    PROC Path_ContornoExterno()
        MoveJ Pivote,v100,z1,MyNewTool\WObj:=Cara;
        MoveJ Target_190,v100,z1,MyNewTool\WObj:=Cara;
        MoveL Target_200,v100,z1,MyNewTool\WObj:=Cara;
        MoveL Target_210,v100,z1,MyNewTool\WObj:=Cara;
        MoveL Target_220,v100,z1,MyNewTool\WObj:=Cara;
        MoveL Target_230,v100,z1,MyNewTool\WObj:=Cara;
        MoveL Target_240,v100,z1,MyNewTool\WObj:=Cara;
        MoveL Target_250,v100,z1,MyNewTool\WObj:=Cara;
        MoveL Target_260,v100,z1,MyNewTool\WObj:=Cara;
        MoveL Target_270,v100,z1,MyNewTool\WObj:=Cara;
        MoveL Target_280,v100,z1,MyNewTool\WObj:=Cara;
        MoveL Target_290,v100,z1,MyNewTool\WObj:=Cara;
        MoveL Target_300,v100,z1,MyNewTool\WObj:=Cara;
        MoveL Target_310,v100,z1,MyNewTool\WObj:=Cara;
        MoveL Target_320,v100,z1,MyNewTool\WObj:=Cara;
        MoveL Target_330,v100,z1,MyNewTool\WObj:=Cara;
        MoveL Target_340,v100,z1,MyNewTool\WObj:=Cara;
        MoveL Target_350,v100,z1,MyNewTool\WObj:=Cara;
        MoveL Target_360,v100,z1,MyNewTool\WObj:=Cara;
        MoveL Target_370,v100,z1,MyNewTool\WObj:=Cara;
        MoveL Target_380,v100,z1,MyNewTool\WObj:=Cara;
        MoveL Target_390,v100,z1,MyNewTool\WObj:=Cara;
        MoveL Target_400,v100,z1,MyNewTool\WObj:=Cara;
        MoveL Target_410,v100,z1,MyNewTool\WObj:=Cara;
        MoveL Target_420,v100,z1,MyNewTool\WObj:=Cara;
        MoveL Target_430,v100,z1,MyNewTool\WObj:=Cara;
        MoveL Target_440,v100,z1,MyNewTool\WObj:=Cara;
        MoveL Target_450,v100,z1,MyNewTool\WObj:=Cara;
        MoveL Target_460,v100,z1,MyNewTool\WObj:=Cara;
        MoveL Target_470,v100,z1,MyNewTool\WObj:=Cara;
        MoveL Target_480,v100,z1,MyNewTool\WObj:=Cara;
        MoveL Target_490,v100,z1,MyNewTool\WObj:=Cara;
        MoveL Target_500,v100,z1,MyNewTool\WObj:=Cara;
        MoveL Target_510,v100,z1,MyNewTool\WObj:=Cara;
        MoveL Target_520,v100,z1,MyNewTool\WObj:=Cara;
        MoveL Target_530,v100,z1,MyNewTool\WObj:=Cara;
        MoveL Target_540,v100,z1,MyNewTool\WObj:=Cara;
        MoveL Target_550,v100,z1,MyNewTool\WObj:=Cara;
        MoveL Target_560,v100,z1,MyNewTool\WObj:=Cara;
        MoveL Target_570,v100,z1,MyNewTool\WObj:=Cara;
        MoveL Target_580,v100,z1,MyNewTool\WObj:=Cara;
        MoveL Target_590,v100,z1,MyNewTool\WObj:=Cara;
        MoveL Target_600,v100,z1,MyNewTool\WObj:=Cara;
        MoveL Target_610,v100,z1,MyNewTool\WObj:=Cara;
        MoveL Target_620,v100,z1,MyNewTool\WObj:=Cara;
        MoveL Target_630,v100,z1,MyNewTool\WObj:=Cara;
        MoveL Target_640,v100,z1,MyNewTool\WObj:=Cara;
        MoveL Target_650,v100,z1,MyNewTool\WObj:=Cara;
        MoveL Target_660,v100,z1,MyNewTool\WObj:=Cara;
        MoveL Target_670,v100,z1,MyNewTool\WObj:=Cara;
        MoveL Target_680,v100,z1,MyNewTool\WObj:=Cara;
        MoveL Target_690,v100,z1,MyNewTool\WObj:=Cara;
        MoveL Target_700,v100,z1,MyNewTool\WObj:=Cara;
        MoveL Target_710,v100,z1,MyNewTool\WObj:=Cara;
        MoveL Target_720,v100,z1,MyNewTool\WObj:=Cara;
        MoveL Target_730,v100,z1,MyNewTool\WObj:=Cara;
        MoveL Target_740,v100,z1,MyNewTool\WObj:=Cara;
        MoveL Target_750,v100,z1,MyNewTool\WObj:=Cara;
        MoveL Target_760,v100,z1,MyNewTool\WObj:=Cara;
        MoveL Target_770,v100,z1,MyNewTool\WObj:=Cara;
        MoveL Target_780,v100,z1,MyNewTool\WObj:=Cara;
        MoveL Target_790,v100,z1,MyNewTool\WObj:=Cara;
        MoveL Target_800,v100,z1,MyNewTool\WObj:=Cara;
        MoveL Target_810,v100,z1,MyNewTool\WObj:=Cara;
        MoveL Target_820,v100,z1,MyNewTool\WObj:=Cara;
        MoveL Target_830,v100,z1,MyNewTool\WObj:=Cara;
        MoveL Target_840,v100,z1,MyNewTool\WObj:=Cara;
        MoveL Target_850,v100,z1,MyNewTool\WObj:=Cara;
        MoveL Target_860,v100,z1,MyNewTool\WObj:=Cara;
        MoveL Target_870,v100,z1,MyNewTool\WObj:=Cara;
        MoveL Target_880,v100,z1,MyNewTool\WObj:=Cara;
        MoveL Target_890,v100,z1,MyNewTool\WObj:=Cara;
        MoveL Target_900,v100,z1,MyNewTool\WObj:=Cara;
        MoveL Target_910,v100,z1,MyNewTool\WObj:=Cara;
        MoveL Target_920,v100,z1,MyNewTool\WObj:=Cara;
        MoveL Target_930,v100,z1,MyNewTool\WObj:=Cara;
        MoveL Target_940,v100,z1,MyNewTool\WObj:=Cara;
        MoveL Target_950,v100,z1,MyNewTool\WObj:=Cara;
        MoveL Target_960,v100,z1,MyNewTool\WObj:=Cara;
        MoveL Target_970,v100,z1,MyNewTool\WObj:=Cara;
        MoveL Target_980,v100,z1,MyNewTool\WObj:=Cara;
        MoveL Target_990,v100,z1,MyNewTool\WObj:=Cara;
        MoveL Target_1000,v100,z1,MyNewTool\WObj:=Cara;
        MoveL Target_1010,v100,z1,MyNewTool\WObj:=Cara;
        MoveL Target_1020,v100,z1,MyNewTool\WObj:=Cara;
        MoveL Target_1030,v100,z1,MyNewTool\WObj:=Cara;
        MoveL Target_1040,v100,z1,MyNewTool\WObj:=Cara;
        MoveL Target_1050,v100,z1,MyNewTool\WObj:=Cara;
        MoveL Target_1060,v100,z1,MyNewTool\WObj:=Cara;
        MoveL Target_1070,v100,z1,MyNewTool\WObj:=Cara;
        MoveL Target_1080,v100,z1,MyNewTool\WObj:=Cara;
        MoveL Target_1090,v100,z1,MyNewTool\WObj:=Cara;
        MoveL Target_1100,v100,z1,MyNewTool\WObj:=Cara;
        MoveL Target_1110,v100,z1,MyNewTool\WObj:=Cara;
        MoveL Target_1120,v100,z1,MyNewTool\WObj:=Cara;
        MoveL Target_1130,v100,z1,MyNewTool\WObj:=Cara;
        MoveL Target_1140,v100,z1,MyNewTool\WObj:=Cara;
        MoveL Target_1150,v100,z1,MyNewTool\WObj:=Cara;
        MoveL Target_1160,v100,z1,MyNewTool\WObj:=Cara;
        MoveL Target_1170,v100,z1,MyNewTool\WObj:=Cara;
    ENDPROC
    PROC Path_Cabello()
        MoveJ Target_1350,v100,z1,MyNewTool\WObj:=Cara;
        MoveL Target_1360,v100,z1,MyNewTool\WObj:=Cara;
        MoveL Target_1370,v100,z1,MyNewTool\WObj:=Cara;
        MoveL Target_1380,v100,z1,MyNewTool\WObj:=Cara;
        MoveL Target_1390,v100,z1,MyNewTool\WObj:=Cara;
        MoveL Target_1400,v100,z1,MyNewTool\WObj:=Cara;
        MoveL Target_1410,v100,z1,MyNewTool\WObj:=Cara;
        MoveL Target_1420,v100,z1,MyNewTool\WObj:=Cara;
        MoveL Target_1430,v100,z1,MyNewTool\WObj:=Cara;
        MoveL Target_1440,v100,z1,MyNewTool\WObj:=Cara;
        MoveL Target_1450,v100,z1,MyNewTool\WObj:=Cara;
        MoveL Target_1460,v100,z1,MyNewTool\WObj:=Cara;
        MoveL Target_1470,v100,z1,MyNewTool\WObj:=Cara;
        MoveL Target_1480,v100,z1,MyNewTool\WObj:=Cara;
        MoveL Target_1490,v100,z1,MyNewTool\WObj:=Cara;
        MoveL Target_1500,v100,z1,MyNewTool\WObj:=Cara;
        MoveL Target_1510,v100,z1,MyNewTool\WObj:=Cara;
        MoveL Target_1520,v100,z1,MyNewTool\WObj:=Cara;
        MoveL Target_1530,v100,z1,MyNewTool\WObj:=Cara;
        MoveL Target_1540,v100,z1,MyNewTool\WObj:=Cara;
        MoveL Target_1550,v100,z1,MyNewTool\WObj:=Cara;
        MoveL Target_1560,v100,z1,MyNewTool\WObj:=Cara;
        MoveL Target_1570,v100,z1,MyNewTool\WObj:=Cara;
        MoveL Target_1580,v100,z1,MyNewTool\WObj:=Cara;
        MoveL Target_1590,v100,z1,MyNewTool\WObj:=Cara;
        MoveL Target_1600,v100,z1,MyNewTool\WObj:=Cara;
        MoveL Target_1610,v100,z1,MyNewTool\WObj:=Cara;
        MoveL Target_1620,v100,z1,MyNewTool\WObj:=Cara;
        MoveL Target_1630,v100,z1,MyNewTool\WObj:=Cara;
        MoveL Target_1640,v100,z1,MyNewTool\WObj:=Cara;
        MoveL Target_1650,v100,z1,MyNewTool\WObj:=Cara;
        MoveL Target_1660,v100,z1,MyNewTool\WObj:=Cara;
        MoveL Target_1670,v100,z1,MyNewTool\WObj:=Cara;
        MoveL Target_1680,v100,z1,MyNewTool\WObj:=Cara;
        MoveL Target_1690,v100,z1,MyNewTool\WObj:=Cara;
        MoveL Target_1700,v100,z1,MyNewTool\WObj:=Cara;
        MoveL Target_1710,v100,z1,MyNewTool\WObj:=Cara;
        MoveL Target_1720,v100,z1,MyNewTool\WObj:=Cara;
        MoveL Target_1730,v100,z1,MyNewTool\WObj:=Cara;
        MoveL Target_1740,v100,z1,MyNewTool\WObj:=Cara;
        MoveL Target_1750,v100,z1,MyNewTool\WObj:=Cara;
        MoveL Target_1760,v100,z1,MyNewTool\WObj:=Cara;
        MoveL Target_1770,v100,z1,MyNewTool\WObj:=Cara;
        MoveL Target_1780,v100,z1,MyNewTool\WObj:=Cara;
        MoveL Target_1790,v100,z1,MyNewTool\WObj:=Cara;
        MoveL Target_1800,v100,z1,MyNewTool\WObj:=Cara;
        MoveL Target_1810,v100,z1,MyNewTool\WObj:=Cara;
        MoveL Target_1820,v100,z1,MyNewTool\WObj:=Cara;
        MoveL Target_1830,v100,z1,MyNewTool\WObj:=Cara;
        MoveL Target_1840,v100,z1,MyNewTool\WObj:=Cara;
        MoveL Target_1850,v100,z1,MyNewTool\WObj:=Cara;
        MoveL Target_1860,v100,z1,MyNewTool\WObj:=Cara;
        MoveL Target_1870,v100,z1,MyNewTool\WObj:=Cara;
        MoveL Target_1880,v100,z1,MyNewTool\WObj:=Cara;
        MoveL Target_1890,v100,z1,MyNewTool\WObj:=Cara;
        MoveL Target_1900,v100,z1,MyNewTool\WObj:=Cara;
        MoveL Target_1910,v100,z1,MyNewTool\WObj:=Cara;
        MoveL Target_1920,v100,z1,MyNewTool\WObj:=Cara;
        MoveL Target_1930,v100,z1,MyNewTool\WObj:=Cara;
        MoveL Target_1940,v100,z1,MyNewTool\WObj:=Cara;
        MoveL Target_1950,v100,z1,MyNewTool\WObj:=Cara;
        MoveL Target_1960,v100,z1,MyNewTool\WObj:=Cara;
        MoveL Target_1970,v100,z1,MyNewTool\WObj:=Cara;
        MoveL Target_1980,v100,z1,MyNewTool\WObj:=Cara;
        MoveL Target_1990,v100,z1,MyNewTool\WObj:=Cara;
        MoveL Target_2000,v100,z1,MyNewTool\WObj:=Cara;
        MoveL Target_2010,v100,z1,MyNewTool\WObj:=Cara;
        MoveL Target_2020,v100,z1,MyNewTool\WObj:=Cara;
        MoveL Target_2030,v100,z1,MyNewTool\WObj:=Cara;
        MoveL Target_2040,v100,z1,MyNewTool\WObj:=Cara;
        MoveL Target_2050,v100,z1,MyNewTool\WObj:=Cara;
        MoveL Target_2060,v100,z1,MyNewTool\WObj:=Cara;
        MoveL Target_2070,v100,z1,MyNewTool\WObj:=Cara;
        MoveL Target_2080,v100,z1,MyNewTool\WObj:=Cara;
        MoveL Target_2090,v100,z1,MyNewTool\WObj:=Cara;
        MoveL Target_2100,v100,z1,MyNewTool\WObj:=Cara;
        MoveL Target_2110,v100,z1,MyNewTool\WObj:=Cara;
        MoveL Target_2120,v100,z1,MyNewTool\WObj:=Cara;
        MoveL Target_2130,v100,z1,MyNewTool\WObj:=Cara;
        MoveL Target_2140,v100,z1,MyNewTool\WObj:=Cara;
        MoveL Target_2150,v100,z1,MyNewTool\WObj:=Cara;
    ENDPROC
    PROC Path_Frente()
        MoveJ Target_2430,v100,z1,MyNewTool\WObj:=Cara;
        MoveL Target_2440,v100,z1,MyNewTool\WObj:=Cara;
        MoveL Target_2450,v100,z1,MyNewTool\WObj:=Cara;
        MoveL Target_2460,v100,z1,MyNewTool\WObj:=Cara;
        MoveL Target_2470,v100,z1,MyNewTool\WObj:=Cara;
        MoveL Target_2480,v100,z1,MyNewTool\WObj:=Cara;
        MoveL Target_2490,v100,z1,MyNewTool\WObj:=Cara;
        MoveL Target_2500,v100,z1,MyNewTool\WObj:=Cara;
        MoveL Target_2510,v100,z1,MyNewTool\WObj:=Cara;
        MoveL Target_2520,v100,z1,MyNewTool\WObj:=Cara;
        MoveL Target_2530,v100,z1,MyNewTool\WObj:=Cara;
        MoveL Target_2540,v100,z1,MyNewTool\WObj:=Cara;
        MoveL Target_2550,v100,z1,MyNewTool\WObj:=Cara;
        MoveL Target_2560,v100,z1,MyNewTool\WObj:=Cara;
        MoveL Target_2570,v100,z1,MyNewTool\WObj:=Cara;
        MoveL Target_2580,v100,z1,MyNewTool\WObj:=Cara;
        MoveL Target_2590,v100,z1,MyNewTool\WObj:=Cara;
        MoveL Target_2600,v100,z1,MyNewTool\WObj:=Cara;
        MoveL Target_2610,v100,z1,MyNewTool\WObj:=Cara;
        MoveL Target_2620,v100,z1,MyNewTool\WObj:=Cara;
        MoveL Target_2630,v100,z1,MyNewTool\WObj:=Cara;
        MoveL Target_2640,v100,z1,MyNewTool\WObj:=Cara;
        MoveL Target_2650,v100,z1,MyNewTool\WObj:=Cara;
        MoveL Target_2660,v100,z1,MyNewTool\WObj:=Cara;
        MoveL Target_2670,v100,z1,MyNewTool\WObj:=Cara;
        MoveL Target_2680,v100,z1,MyNewTool\WObj:=Cara;
        MoveL Target_2690,v100,z1,MyNewTool\WObj:=Cara;
        MoveL Target_2700,v100,z1,MyNewTool\WObj:=Cara;
    ENDPROC
    PROC Path_ContornoCara()
        MoveJ Target_2710,v100,z1,MyNewTool\WObj:=Cara;
        MoveL Target_2720,v100,z1,MyNewTool\WObj:=Cara;
        MoveL Target_2730,v100,z1,MyNewTool\WObj:=Cara;
        MoveL Target_2740,v100,z1,MyNewTool\WObj:=Cara;
        MoveL Target_2750,v100,z1,MyNewTool\WObj:=Cara;
        MoveL Target_2760,v100,z1,MyNewTool\WObj:=Cara;
        MoveL Target_2770,v100,z1,MyNewTool\WObj:=Cara;
        MoveL Target_2780,v100,z1,MyNewTool\WObj:=Cara;
        MoveL Target_2790,v100,z1,MyNewTool\WObj:=Cara;
        MoveL Target_2800,v100,z1,MyNewTool\WObj:=Cara;
        MoveL Target_2810,v100,z1,MyNewTool\WObj:=Cara;
        MoveL Target_2820,v100,z1,MyNewTool\WObj:=Cara;
        MoveL Target_2830,v100,z1,MyNewTool\WObj:=Cara;
        MoveL Target_2840,v100,z1,MyNewTool\WObj:=Cara;
        MoveL Target_2850,v100,z1,MyNewTool\WObj:=Cara;
        MoveL Target_2860,v100,z1,MyNewTool\WObj:=Cara;
        MoveL Target_2870,v100,z1,MyNewTool\WObj:=Cara;
        MoveL Target_2880,v100,z1,MyNewTool\WObj:=Cara;
        MoveL Target_2890,v100,z1,MyNewTool\WObj:=Cara;
        MoveL Target_2900,v100,z1,MyNewTool\WObj:=Cara;
        MoveL Target_2910,v100,z1,MyNewTool\WObj:=Cara;
        MoveL Target_2920,v100,z1,MyNewTool\WObj:=Cara;
        MoveL Target_2930,v100,z1,MyNewTool\WObj:=Cara;
        MoveL Target_2940,v100,z1,MyNewTool\WObj:=Cara;
        MoveL Target_2950,v100,z1,MyNewTool\WObj:=Cara;
        MoveL Target_2960,v100,z1,MyNewTool\WObj:=Cara;
        MoveL Target_2970,v100,z1,MyNewTool\WObj:=Cara;
        MoveL Target_2980,v100,z1,MyNewTool\WObj:=Cara;
        MoveL Target_2990,v100,z1,MyNewTool\WObj:=Cara;
        MoveL Target_3000,v100,z1,MyNewTool\WObj:=Cara;
        MoveL Target_3010,v100,z1,MyNewTool\WObj:=Cara;
        MoveL Target_3020,v100,z1,MyNewTool\WObj:=Cara;
        MoveL Target_3030,v100,z1,MyNewTool\WObj:=Cara;
        MoveL Target_3040,v100,z1,MyNewTool\WObj:=Cara;
        MoveL Target_3050,v100,z1,MyNewTool\WObj:=Cara;
        MoveL Target_3060,v100,z1,MyNewTool\WObj:=Cara;
        MoveL Target_3070,v100,z1,MyNewTool\WObj:=Cara;
        MoveL Target_3080,v100,z1,MyNewTool\WObj:=Cara;
        MoveL Target_3090,v100,z1,MyNewTool\WObj:=Cara;
        MoveL Target_3100,v100,z1,MyNewTool\WObj:=Cara;
        MoveL Target_3110,v100,z1,MyNewTool\WObj:=Cara;
        MoveL Target_3120,v100,z1,MyNewTool\WObj:=Cara;
        MoveL Target_3130,v100,z1,MyNewTool\WObj:=Cara;
        MoveL Target_3140,v100,z1,MyNewTool\WObj:=Cara;
        MoveL Target_3150,v100,z1,MyNewTool\WObj:=Cara;
        MoveL Target_3160,v100,z1,MyNewTool\WObj:=Cara;
        MoveL Target_3170,v100,z1,MyNewTool\WObj:=Cara;
        MoveL Target_3180,v100,z1,MyNewTool\WObj:=Cara;
        MoveL Target_3190,v100,z1,MyNewTool\WObj:=Cara;
        MoveL Target_3200,v100,z1,MyNewTool\WObj:=Cara;
        MoveL Target_3210,v100,z1,MyNewTool\WObj:=Cara;
        MoveL Target_3220,v100,z1,MyNewTool\WObj:=Cara;
        MoveL Target_3230,v100,z1,MyNewTool\WObj:=Cara;
        MoveL Target_3240,v100,z1,MyNewTool\WObj:=Cara;
        MoveL Target_3250,v100,z1,MyNewTool\WObj:=Cara;
        MoveL Target_3260,v100,z1,MyNewTool\WObj:=Cara;
        MoveL Target_3270,v100,z1,MyNewTool\WObj:=Cara;
        MoveL Target_3280,v100,z1,MyNewTool\WObj:=Cara;
        MoveL Target_3290,v100,z1,MyNewTool\WObj:=Cara;
        MoveL Target_3300,v100,z1,MyNewTool\WObj:=Cara;
        MoveL Target_3310,v100,z1,MyNewTool\WObj:=Cara;
        MoveL Target_3320,v100,z1,MyNewTool\WObj:=Cara;
        MoveL Target_3330,v100,z1,MyNewTool\WObj:=Cara;
        MoveL Target_3340,v100,z1,MyNewTool\WObj:=Cara;
        MoveL Target_3350,v100,z1,MyNewTool\WObj:=Cara;
        MoveL Target_3360,v100,z1,MyNewTool\WObj:=Cara;
        MoveL Target_3370,v100,z1,MyNewTool\WObj:=Cara;
        MoveL Target_3380,v100,z1,MyNewTool\WObj:=Cara;
        MoveL Target_3390,v100,z1,MyNewTool\WObj:=Cara;
        MoveL Target_3400,v100,z1,MyNewTool\WObj:=Cara;
        MoveL Target_3410,v100,z1,MyNewTool\WObj:=Cara;
        MoveL Target_3420,v100,z1,MyNewTool\WObj:=Cara;
        MoveL Target_3430,v100,z1,MyNewTool\WObj:=Cara;
        MoveL Target_3440,v100,z1,MyNewTool\WObj:=Cara;
        MoveL Target_3450,v100,z1,MyNewTool\WObj:=Cara;
        MoveL Target_3460,v100,z1,MyNewTool\WObj:=Cara;
        MoveL Target_3470,v100,z1,MyNewTool\WObj:=Cara;
        MoveL Target_3480,v100,z1,MyNewTool\WObj:=Cara;
        MoveL Target_3490,v100,z1,MyNewTool\WObj:=Cara;
        MoveL Target_3500,v100,z1,MyNewTool\WObj:=Cara;
        MoveL Target_3510,v100,z1,MyNewTool\WObj:=Cara;
        MoveL Target_3520,v100,z1,MyNewTool\WObj:=Cara;
        MoveL Target_3530,v100,z1,MyNewTool\WObj:=Cara;
        MoveL Target_3540,v100,z1,MyNewTool\WObj:=Cara;
        MoveL Target_3550,v100,z1,MyNewTool\WObj:=Cara;
        MoveL Target_3560,v100,z1,MyNewTool\WObj:=Cara;
        MoveL Target_3570,v100,z1,MyNewTool\WObj:=Cara;
        MoveL Target_3580,v100,z1,MyNewTool\WObj:=Cara;
        MoveL Target_3590,v100,z1,MyNewTool\WObj:=Cara;
        MoveL Target_3600,v100,z1,MyNewTool\WObj:=Cara;
        MoveL Target_3610,v100,z1,MyNewTool\WObj:=Cara;
        MoveL Target_3620,v100,z1,MyNewTool\WObj:=Cara;
        MoveL Target_3630,v100,z1,MyNewTool\WObj:=Cara;
        MoveL Target_3640,v100,z1,MyNewTool\WObj:=Cara;
        MoveL Target_3650,v100,z1,MyNewTool\WObj:=Cara;
        MoveL Target_3660,v100,z1,MyNewTool\WObj:=Cara;
        MoveL Target_3670,v100,z1,MyNewTool\WObj:=Cara;
        MoveL Target_3680,v100,z1,MyNewTool\WObj:=Cara;
        MoveL Target_3690,v100,z1,MyNewTool\WObj:=Cara;
        MoveL Target_3700,v100,z1,MyNewTool\WObj:=Cara;
        MoveL Target_3710,v100,z1,MyNewTool\WObj:=Cara;
    ENDPROC
    PROC Path_Boca()
        MoveJ Target_3720,v100,z1,MyNewTool\WObj:=Cara;
        MoveL Target_3730,v100,z1,MyNewTool\WObj:=Cara;
        MoveL Target_3740,v100,z1,MyNewTool\WObj:=Cara;
        MoveL Target_3750,v100,z1,MyNewTool\WObj:=Cara;
        MoveL Target_3760,v100,z1,MyNewTool\WObj:=Cara;
        MoveL Target_3770,v100,z1,MyNewTool\WObj:=Cara;
        MoveL Target_3780,v100,z1,MyNewTool\WObj:=Cara;
        MoveL Target_3790,v100,z1,MyNewTool\WObj:=Cara;
        MoveL Target_3800,v100,z1,MyNewTool\WObj:=Cara;
        MoveL Target_3810,v100,z1,MyNewTool\WObj:=Cara;
        MoveL Target_3820,v100,z1,MyNewTool\WObj:=Cara;
    ENDPROC
    PROC Path_BandaNinja()
        MoveJ Target_10,v100,z1,MyNewTool\WObj:=Cara;
        MoveL Target_20,v100,z1,MyNewTool\WObj:=Cara;
        MoveL Target_30,v100,z1,MyNewTool\WObj:=Cara;
        MoveL Target_40,v100,z1,MyNewTool\WObj:=Cara;
        MoveL Target_50,v100,z1,MyNewTool\WObj:=Cara;
        MoveL Target_60,v100,z1,MyNewTool\WObj:=Cara;
        MoveL Target_70,v100,z1,MyNewTool\WObj:=Cara;
        MoveL Target_80,v100,z1,MyNewTool\WObj:=Cara;
        MoveL Target_90,v100,z1,MyNewTool\WObj:=Cara;
        MoveL Target_100,v100,z1,MyNewTool\WObj:=Cara;
        MoveL Target_110,v100,z1,MyNewTool\WObj:=Cara;
        MoveL Target_120,v100,z1,MyNewTool\WObj:=Cara;
        MoveL Target_130,v100,z1,MyNewTool\WObj:=Cara;
        MoveL Target_140,v100,z1,MyNewTool\WObj:=Cara;
        MoveL Target_150,v100,z1,MyNewTool\WObj:=Cara;
        MoveL Target_160,v100,z1,MyNewTool\WObj:=Cara;
        MoveL Target_170,v100,z1,MyNewTool\WObj:=Cara;
        MoveL Target_180,v100,z1,MyNewTool\WObj:=Cara;
    ENDPROC
    PROC Path_SimboloNinja()
        MoveJ Target_2160,v100,z1,MyNewTool\WObj:=Cara;
        MoveL Target_2170,v100,z1,MyNewTool\WObj:=Cara;
        MoveL Target_2180,v100,z1,MyNewTool\WObj:=Cara;
        MoveL Target_2190,v100,z1,MyNewTool\WObj:=Cara;
        MoveL Target_2200,v100,z1,MyNewTool\WObj:=Cara;
        MoveL Target_2210,v100,z1,MyNewTool\WObj:=Cara;
        MoveL Target_2220,v100,z1,MyNewTool\WObj:=Cara;
        MoveL Target_2230,v100,z1,MyNewTool\WObj:=Cara;
        MoveL Target_2240,v100,z1,MyNewTool\WObj:=Cara;
        MoveL Target_2250,v100,z1,MyNewTool\WObj:=Cara;
        MoveL Target_2260,v100,z1,MyNewTool\WObj:=Cara;
        MoveL Target_2270,v100,z1,MyNewTool\WObj:=Cara;
        MoveL Target_2280,v100,z1,MyNewTool\WObj:=Cara;
        MoveL Target_2290,v100,z1,MyNewTool\WObj:=Cara;
        MoveL Target_2300,v100,z1,MyNewTool\WObj:=Cara;
        MoveL Target_2310,v100,z1,MyNewTool\WObj:=Cara;
        MoveL Target_2320,v100,z1,MyNewTool\WObj:=Cara;
        MoveL Target_2330,v100,z1,MyNewTool\WObj:=Cara;
        MoveL Target_2340,v100,z1,MyNewTool\WObj:=Cara;
        MoveL Target_2350,v100,z1,MyNewTool\WObj:=Cara;
        MoveL Target_2360,v100,z1,MyNewTool\WObj:=Cara;
        MoveL Target_2370,v100,z1,MyNewTool\WObj:=Cara;
        MoveL Target_2380,v100,z1,MyNewTool\WObj:=Cara;
        MoveL Target_2390,v100,z1,MyNewTool\WObj:=Cara;
        MoveL Target_2400,v100,z1,MyNewTool\WObj:=Cara;
        MoveL Target_2410,v100,z1,MyNewTool\WObj:=Cara;
        MoveL Target_2420,v100,z1,MyNewTool\WObj:=Cara;
    ENDPROC
    PROC Path_OrejaDerecha1()
        MoveJ Target_3830,v100,z1,MyNewTool\WObj:=Cara;
        MoveL Target_3840,v100,z1,MyNewTool\WObj:=Cara;
        MoveL Target_3850,v100,z1,MyNewTool\WObj:=Cara;
        MoveL Target_3860,v100,z1,MyNewTool\WObj:=Cara;
        MoveL Target_3870,v100,z1,MyNewTool\WObj:=Cara;
        MoveL Target_3880,v100,z1,MyNewTool\WObj:=Cara;
        MoveL Target_3890,v100,z1,MyNewTool\WObj:=Cara;
        MoveL Target_3900,v100,z1,MyNewTool\WObj:=Cara;
        MoveL Target_3910,v100,z1,MyNewTool\WObj:=Cara;
        MoveL Target_3920,v100,z1,MyNewTool\WObj:=Cara;
        MoveL Target_3930,v100,z1,MyNewTool\WObj:=Cara;
        MoveL Target_3940,v100,z1,MyNewTool\WObj:=Cara;
        MoveL Target_3950,v100,z1,MyNewTool\WObj:=Cara;
        MoveL Target_3960,v100,z1,MyNewTool\WObj:=Cara;
        MoveL Target_3970,v100,z1,MyNewTool\WObj:=Cara;
        MoveL Target_3980,v100,z1,MyNewTool\WObj:=Cara;
        MoveL Target_3990,v100,z1,MyNewTool\WObj:=Cara;
    ENDPROC
    PROC Path_OrejaDerecha2()
        MoveJ Target_4000,v100,z1,MyNewTool\WObj:=Cara;
        MoveL Target_4010,v100,z1,MyNewTool\WObj:=Cara;
        MoveL Target_4020,v100,z1,MyNewTool\WObj:=Cara;
        MoveL Target_4030,v100,z1,MyNewTool\WObj:=Cara;
        MoveL Target_4040,v100,z1,MyNewTool\WObj:=Cara;
        MoveL Target_4050,v100,z1,MyNewTool\WObj:=Cara;
        MoveL Target_4060,v100,z1,MyNewTool\WObj:=Cara;
        MoveL Target_4070,v100,z1,MyNewTool\WObj:=Cara;
        MoveL Target_4080,v100,z1,MyNewTool\WObj:=Cara;
        MoveL Target_4090,v100,z1,MyNewTool\WObj:=Cara;
    ENDPROC
    PROC Path_OrejaIzquierda2()
        MoveJ Target_4100,v100,z1,MyNewTool\WObj:=Cara;
        MoveL Target_4110,v100,z1,MyNewTool\WObj:=Cara;
        MoveL Target_4120,v100,z1,MyNewTool\WObj:=Cara;
        MoveL Target_4130,v100,z1,MyNewTool\WObj:=Cara;
        MoveL Target_4140,v100,z1,MyNewTool\WObj:=Cara;
        MoveL Target_4150,v100,z1,MyNewTool\WObj:=Cara;
        MoveL Target_4160,v100,z1,MyNewTool\WObj:=Cara;
        MoveL Target_4170,v100,z1,MyNewTool\WObj:=Cara;
        MoveL Target_4180,v100,z1,MyNewTool\WObj:=Cara;
        MoveL Target_4190,v100,z1,MyNewTool\WObj:=Cara;
    ENDPROC
    PROC Path_OrejaIzquierda1()
        MoveJ Target_4200,v100,z1,MyNewTool\WObj:=Cara;
        MoveL Target_4210,v100,z1,MyNewTool\WObj:=Cara;
        MoveL Target_4220,v100,z1,MyNewTool\WObj:=Cara;
        MoveL Target_4230,v100,z1,MyNewTool\WObj:=Cara;
        MoveL Target_4240,v100,z1,MyNewTool\WObj:=Cara;
        MoveL Target_4250,v100,z1,MyNewTool\WObj:=Cara;
        MoveL Target_4260,v100,z1,MyNewTool\WObj:=Cara;
        MoveL Target_4270,v100,z1,MyNewTool\WObj:=Cara;
        MoveL Target_4280,v100,z1,MyNewTool\WObj:=Cara;
        MoveL Target_4290,v100,z1,MyNewTool\WObj:=Cara;
        MoveL Target_4300,v100,z1,MyNewTool\WObj:=Cara;
        MoveL Target_4310,v100,z1,MyNewTool\WObj:=Cara;
        MoveL Target_4320,v100,z1,MyNewTool\WObj:=Cara;
        MoveL Target_4330,v100,z1,MyNewTool\WObj:=Cara;
        MoveL Target_4340,v100,z1,MyNewTool\WObj:=Cara;
        MoveL Target_4350,v100,z1,MyNewTool\WObj:=Cara;
    ENDPROC
    PROC Path_Detalle1()
        MoveJ Target_4490,v100,z1,MyNewTool\WObj:=Cara;
        MoveL Target_4500,v100,z1,MyNewTool\WObj:=Cara;
        MoveL Target_4510,v100,z1,MyNewTool\WObj:=Cara;
    ENDPROC
    PROC Path_Detalle2()
        MoveJ Target_4520,v100,z1,MyNewTool\WObj:=Cara;
        MoveL Target_4530,v100,z1,MyNewTool\WObj:=Cara;
        MoveL Target_4540,v100,z1,MyNewTool\WObj:=Cara;
    ENDPROC
    PROC Path_Detalle3()
        MoveJ Target_4550,v100,z1,MyNewTool\WObj:=Cara;
        MoveL Target_4560,v100,z1,MyNewTool\WObj:=Cara;
        MoveL Target_4570,v100,z1,MyNewTool\WObj:=Cara;
    ENDPROC
    PROC Path_Pintar1()
        MoveJ Target_4580,v100,z1,MyNewTool\WObj:=Cara;
        MoveL Target_4590,v100,z1,MyNewTool\WObj:=Cara;
        MoveL Target_4600,v100,z1,MyNewTool\WObj:=Cara;
        MoveL Target_4610,v100,z1,MyNewTool\WObj:=Cara;
        MoveL Target_4620,v100,z1,MyNewTool\WObj:=Cara;
        MoveL Target_4630,v100,z1,MyNewTool\WObj:=Cara;
        MoveL Target_4640,v100,z1,MyNewTool\WObj:=Cara;
        MoveL Target_4650,v100,z1,MyNewTool\WObj:=Cara;
        MoveL Target_4660,v100,z1,MyNewTool\WObj:=Cara;
        MoveL Target_4670,v100,z1,MyNewTool\WObj:=Cara;
        MoveL Target_4680,v100,z1,MyNewTool\WObj:=Cara;
        MoveL Target_4690,v100,z1,MyNewTool\WObj:=Cara;
        MoveL Target_4700,v100,z1,MyNewTool\WObj:=Cara;
        MoveL Target_4710,v100,z1,MyNewTool\WObj:=Cara;
        MoveL Target_4720,v100,z1,MyNewTool\WObj:=Cara;
        MoveL Target_4730,v100,z1,MyNewTool\WObj:=Cara;
        MoveL Target_4740,v100,z1,MyNewTool\WObj:=Cara;
        MoveL Target_4750,v100,z1,MyNewTool\WObj:=Cara;
    ENDPROC
    PROC Path_Detalle5()
        MoveJ Target_4760,v100,z1,MyNewTool\WObj:=Cara;
        MoveL Target_4770,v100,z1,MyNewTool\WObj:=Cara;
        MoveL Target_4780,v100,z1,MyNewTool\WObj:=Cara;
        MoveL Target_4790,v100,z1,MyNewTool\WObj:=Cara;
        MoveL Target_4800,v100,z1,MyNewTool\WObj:=Cara;
    ENDPROC
    PROC Path_Detalle4()
        MoveJ Target_4810,v100,z1,MyNewTool\WObj:=Cara;
        MoveL Target_4820,v100,z1,MyNewTool\WObj:=Cara;
        MoveL Target_4830,v100,z1,MyNewTool\WObj:=Cara;
        MoveL Target_4840,v100,z1,MyNewTool\WObj:=Cara;
        MoveL Target_4850,v100,z1,MyNewTool\WObj:=Cara;
    ENDPROC
    PROC Path_Pintar2()
        MoveJ Target_4860,v100,z1,MyNewTool\WObj:=Cara;
        MoveL Target_4870,v100,z1,MyNewTool\WObj:=Cara;
        MoveL Target_4880,v100,z1,MyNewTool\WObj:=Cara;
        MoveL Target_4890,v100,z1,MyNewTool\WObj:=Cara;
        MoveL Target_4900,v100,z1,MyNewTool\WObj:=Cara;
        MoveL Target_4910,v100,z1,MyNewTool\WObj:=Cara;
        MoveL Target_4920,v100,z1,MyNewTool\WObj:=Cara;
        MoveL Target_4930,v100,z1,MyNewTool\WObj:=Cara;
        MoveL Target_4940,v100,z1,MyNewTool\WObj:=Cara;
        MoveL Target_4950,v100,z1,MyNewTool\WObj:=Cara;
        MoveL Target_4960,v100,z1,MyNewTool\WObj:=Cara;
        MoveL Target_4970,v100,z1,MyNewTool\WObj:=Cara;
        MoveL Target_4980,v100,z1,MyNewTool\WObj:=Cara;
        MoveL Target_4990,v100,z1,MyNewTool\WObj:=Cara;
        MoveL Target_5000,v100,z1,MyNewTool\WObj:=Cara;
        MoveL Target_5010,v100,z1,MyNewTool\WObj:=Cara;
        MoveL Target_5020,v100,z1,MyNewTool\WObj:=Cara;
        MoveL Target_5030,v100,z1,MyNewTool\WObj:=Cara;
        MoveL Target_5040,v100,z1,MyNewTool\WObj:=Cara;
        MoveL Target_5050,v100,z1,MyNewTool\WObj:=Cara;
        MoveL Target_5060,v100,z1,MyNewTool\WObj:=Cara;
        MoveL Target_5070,v100,z1,MyNewTool\WObj:=Cara;
        MoveL Target_5080,v100,z1,MyNewTool\WObj:=Cara;
    ENDPROC
    PROC Path_Detalle6()
        MoveJ Target_5090,v100,z1,MyNewTool\WObj:=Cara;
        MoveL Target_5100,v100,z1,MyNewTool\WObj:=Cara;
        MoveL Target_5110,v100,z1,MyNewTool\WObj:=Cara;
        MoveL Target_5120,v100,z1,MyNewTool\WObj:=Cara;
        MoveL Target_5130,v100,z1,MyNewTool\WObj:=Cara;
    ENDPROC
    PROC Path_Detalle7()
        MoveJ Target_5140,v100,z1,MyNewTool\WObj:=Cara;
        MoveL Target_5150,v100,z1,MyNewTool\WObj:=Cara;
        MoveL Target_5160,v100,z1,MyNewTool\WObj:=Cara;
        MoveL Target_5170,v100,z1,MyNewTool\WObj:=Cara;
    ENDPROC
    PROC Path_Home()
        MoveJ Target_Home,v100,fine,MyNewTool\WObj:=Cara;
    ENDPROC
    PROC Path_Pausa()
        MoveJ Target_Pausa,v200,z1,MyNewTool\WObj:=Cara;
    ENDPROC
    PROC Path_Nombre1_A1()
        MoveL Target_5180,v100,z1,MyNewTool\WObj:=Cara;
        MoveL Target_5190,v100,z1,MyNewTool\WObj:=Cara;
        MoveL Target_5200,v100,z1,MyNewTool\WObj:=Cara;
        MoveL Target_5210,v100,z1,MyNewTool\WObj:=Cara;
        MoveL Target_5220,v100,z1,MyNewTool\WObj:=Cara;
        MoveL Target_5230,v100,z1,MyNewTool\WObj:=Cara;
        MoveL Target_5240,v100,z1,MyNewTool\WObj:=Cara;
        MoveL Target_5250,v100,z1,MyNewTool\WObj:=Cara;
        MoveL Target_5260,v100,z1,MyNewTool\WObj:=Cara;
    ENDPROC
    PROC Path_Nombre1_A2()
        MoveL Target_5270,v100,z1,MyNewTool\WObj:=Cara;
        MoveL Target_5280,v100,z1,MyNewTool\WObj:=Cara;
        MoveL Target_5290,v100,z1,MyNewTool\WObj:=Cara;
        MoveL Target_5300,v100,z1,MyNewTool\WObj:=Cara;
    ENDPROC
    PROC Path_Nombre1_R1()
        MoveL Target_5310,v100,z1,MyNewTool\WObj:=Cara;
        MoveL Target_5320,v100,z1,MyNewTool\WObj:=Cara;
        MoveL Target_5330,v100,z1,MyNewTool\WObj:=Cara;
        MoveL Target_5340,v100,z1,MyNewTool\WObj:=Cara;
        MoveL Target_5350,v100,z1,MyNewTool\WObj:=Cara;
        MoveL Target_5360,v100,z1,MyNewTool\WObj:=Cara;
        MoveL Target_5370,v100,z1,MyNewTool\WObj:=Cara;
        MoveL Target_5380,v100,z1,MyNewTool\WObj:=Cara;
        MoveL Target_5390,v100,z1,MyNewTool\WObj:=Cara;
        MoveL Target_5400,v100,z1,MyNewTool\WObj:=Cara;
        MoveL Target_5410,v100,z1,MyNewTool\WObj:=Cara;
        MoveL Target_5420,v100,z1,MyNewTool\WObj:=Cara;
        MoveL Target_5430,v100,z1,MyNewTool\WObj:=Cara;
    ENDPROC
    PROC Path_Nombre1_R2()
        MoveL Target_5440,v100,z1,MyNewTool\WObj:=Cara;
        MoveL Target_5450,v100,z1,MyNewTool\WObj:=Cara;
        MoveL Target_5460,v100,z1,MyNewTool\WObj:=Cara;
        MoveL Target_5470,v100,z1,MyNewTool\WObj:=Cara;
        MoveL Target_5480,v100,z1,MyNewTool\WObj:=Cara;
        MoveL Target_5490,v100,z1,MyNewTool\WObj:=Cara;
    ENDPROC
    PROC Path_Nombre1_I()
        MoveL Target_5500,v100,z1,MyNewTool\WObj:=Cara;
        MoveL Target_5510,v100,z1,MyNewTool\WObj:=Cara;
        MoveL Target_5520,v100,z1,MyNewTool\WObj:=Cara;
        MoveL Target_5530,v100,z1,MyNewTool\WObj:=Cara;
        MoveL Target_5540,v100,z1,MyNewTool\WObj:=Cara;
        MoveL Target_5550,v100,z1,MyNewTool\WObj:=Cara;
        MoveL Target_5560,v100,z1,MyNewTool\WObj:=Cara;
        MoveL Target_5570,v100,z1,MyNewTool\WObj:=Cara;
        MoveL Target_5580,v100,z1,MyNewTool\WObj:=Cara;
        MoveL Target_5590,v100,z1,MyNewTool\WObj:=Cara;
        MoveL Target_5600,v100,z1,MyNewTool\WObj:=Cara;
        MoveL Target_5610,v100,z1,MyNewTool\WObj:=Cara;
        MoveL Target_5620,v100,z1,MyNewTool\WObj:=Cara;
    ENDPROC
    PROC Path_Nombre1_E()
        MoveL Target_5630,v100,z1,MyNewTool\WObj:=Cara;
        MoveL Target_5640,v100,z1,MyNewTool\WObj:=Cara;
        MoveL Target_5650,v100,z1,MyNewTool\WObj:=Cara;
        MoveL Target_5660,v100,z1,MyNewTool\WObj:=Cara;
        MoveL Target_5670,v100,z1,MyNewTool\WObj:=Cara;
        MoveL Target_5680,v100,z1,MyNewTool\WObj:=Cara;
        MoveL Target_5690,v100,z1,MyNewTool\WObj:=Cara;
        MoveL Target_5700,v100,z1,MyNewTool\WObj:=Cara;
        MoveL Target_5710,v100,z1,MyNewTool\WObj:=Cara;
        MoveL Target_5720,v100,z1,MyNewTool\WObj:=Cara;
        MoveL Target_5730,v100,z1,MyNewTool\WObj:=Cara;
        MoveL Target_5740,v100,z1,MyNewTool\WObj:=Cara;
        MoveL Target_5750,v100,z1,MyNewTool\WObj:=Cara;
    ENDPROC
    PROC Path_Nombre1_L()
        MoveL Target_5760,v100,z1,MyNewTool\WObj:=Cara;
        MoveL Target_5770,v100,z1,MyNewTool\WObj:=Cara;
        MoveL Target_5780,v100,z1,MyNewTool\WObj:=Cara;
        MoveL Target_5790,v100,z1,MyNewTool\WObj:=Cara;
        MoveL Target_5800,v100,z1,MyNewTool\WObj:=Cara;
        MoveL Target_5810,v100,z1,MyNewTool\WObj:=Cara;
        MoveL Target_5820,v100,z1,MyNewTool\WObj:=Cara;
    ENDPROC
    PROC Path_Nombre2_J()
        MoveL Target_5830,v100,z1,MyNewTool\WObj:=Cara;
        MoveL Target_5840,v100,z1,MyNewTool\WObj:=Cara;
        MoveL Target_5850,v100,z1,MyNewTool\WObj:=Cara;
        MoveL Target_5860,v100,z1,MyNewTool\WObj:=Cara;
        MoveL Target_5870,v100,z1,MyNewTool\WObj:=Cara;
        MoveL Target_5880,v100,z1,MyNewTool\WObj:=Cara;
        MoveL Target_5890,v100,z1,MyNewTool\WObj:=Cara;
        MoveL Target_5900,v100,z1,MyNewTool\WObj:=Cara;
        MoveL Target_5910,v100,z1,MyNewTool\WObj:=Cara;
        MoveL Target_5920,v100,z1,MyNewTool\WObj:=Cara;
        MoveL Target_5930,v100,z1,MyNewTool\WObj:=Cara;
        MoveL Target_5940,v100,z1,MyNewTool\WObj:=Cara;
    ENDPROC
    PROC Path_Nombre2_A1()
        MoveL Target_5950,v100,z1,MyNewTool\WObj:=Cara;
        MoveL Target_5960,v100,z1,MyNewTool\WObj:=Cara;
        MoveL Target_5970,v100,z1,MyNewTool\WObj:=Cara;
        MoveL Target_5980,v100,z1,MyNewTool\WObj:=Cara;
        MoveL Target_5990,v100,z1,MyNewTool\WObj:=Cara;
        MoveL Target_6000,v100,z1,MyNewTool\WObj:=Cara;
        MoveL Target_6010,v100,z1,MyNewTool\WObj:=Cara;
        MoveL Target_6020,v100,z1,MyNewTool\WObj:=Cara;
        MoveL Target_6030,v100,z1,MyNewTool\WObj:=Cara;
    ENDPROC
    PROC Path_Nombre2_A2()
        MoveL Target_6040,v100,z1,MyNewTool\WObj:=Cara;
        MoveL Target_6050,v100,z1,MyNewTool\WObj:=Cara;
        MoveL Target_6060,v100,z1,MyNewTool\WObj:=Cara;
        MoveL Target_6070,v100,z1,MyNewTool\WObj:=Cara;
    ENDPROC
    PROC Path_Nombre2_R1()
        MoveL Target_6080,v100,z1,MyNewTool\WObj:=Cara;
        MoveL Target_6090,v100,z1,MyNewTool\WObj:=Cara;
        MoveL Target_6100,v100,z1,MyNewTool\WObj:=Cara;
        MoveL Target_6110,v100,z1,MyNewTool\WObj:=Cara;
        MoveL Target_6120,v100,z1,MyNewTool\WObj:=Cara;
        MoveL Target_6130,v100,z1,MyNewTool\WObj:=Cara;
        MoveL Target_6140,v100,z1,MyNewTool\WObj:=Cara;
        MoveL Target_6150,v100,z1,MyNewTool\WObj:=Cara;
        MoveL Target_6160,v100,z1,MyNewTool\WObj:=Cara;
        MoveL Target_6170,v100,z1,MyNewTool\WObj:=Cara;
        MoveL Target_6180,v100,z1,MyNewTool\WObj:=Cara;
        MoveL Target_6190,v100,z1,MyNewTool\WObj:=Cara;
        MoveL Target_6200,v100,z1,MyNewTool\WObj:=Cara;
    ENDPROC
    PROC Path_Nombre2_R2()
        MoveL Target_6210,v100,z1,MyNewTool\WObj:=Cara;
        MoveL Target_6220,v100,z1,MyNewTool\WObj:=Cara;
        MoveL Target_6230,v100,z1,MyNewTool\WObj:=Cara;
        MoveL Target_6240,v100,z1,MyNewTool\WObj:=Cara;
        MoveL Target_6250,v100,z1,MyNewTool\WObj:=Cara;
        MoveL Target_6260,v100,z1,MyNewTool\WObj:=Cara;
    ENDPROC
    PROC Path_Nombre2_E()
        MoveL Target_6270,v100,z1,MyNewTool\WObj:=Cara;
        MoveL Target_6280,v100,z1,MyNewTool\WObj:=Cara;
        MoveL Target_6290,v100,z1,MyNewTool\WObj:=Cara;
        MoveL Target_6300,v100,z1,MyNewTool\WObj:=Cara;
        MoveL Target_6310,v100,z1,MyNewTool\WObj:=Cara;
        MoveL Target_6320,v100,z1,MyNewTool\WObj:=Cara;
        MoveL Target_6330,v100,z1,MyNewTool\WObj:=Cara;
        MoveL Target_6340,v100,z1,MyNewTool\WObj:=Cara;
        MoveL Target_6350,v100,z1,MyNewTool\WObj:=Cara;
        MoveL Target_6360,v100,z1,MyNewTool\WObj:=Cara;
        MoveL Target_6370,v100,z1,MyNewTool\WObj:=Cara;
        MoveL Target_6380,v100,z1,MyNewTool\WObj:=Cara;
        MoveL Target_6390,v100,z1,MyNewTool\WObj:=Cara;
    ENDPROC
    PROC Path_Nombre2_D1()
        MoveL Target_6400,v100,z1,MyNewTool\WObj:=Cara;
        MoveL Target_6410,v100,z1,MyNewTool\WObj:=Cara;
        MoveL Target_6420,v100,z1,MyNewTool\WObj:=Cara;
        MoveL Target_6430,v100,z1,MyNewTool\WObj:=Cara;
        MoveL Target_6440,v100,z1,MyNewTool\WObj:=Cara;
        MoveL Target_6450,v100,z1,MyNewTool\WObj:=Cara;
        MoveL Target_6460,v100,z1,MyNewTool\WObj:=Cara;
        MoveL Target_6470,v100,z1,MyNewTool\WObj:=Cara;
        MoveL Target_6480,v100,z1,MyNewTool\WObj:=Cara;
        MoveL Target_6490,v100,z1,MyNewTool\WObj:=Cara;
        MoveL Target_6500,v100,z1,MyNewTool\WObj:=Cara;
    ENDPROC
    PROC Path_Nombre2_D2()
        MoveL Target_6510,v100,z1,MyNewTool\WObj:=Cara;
        MoveL Target_6520,v100,z1,MyNewTool\WObj:=Cara;
        MoveL Target_6530,v100,z1,MyNewTool\WObj:=Cara;
        MoveL Target_6540,v100,z1,MyNewTool\WObj:=Cara;
        MoveL Target_6550,v100,z1,MyNewTool\WObj:=Cara;
        MoveL Target_6560,v100,z1,MyNewTool\WObj:=Cara;
        MoveL Target_6570,v100,z1,MyNewTool\WObj:=Cara;
        MoveL Target_6580,v100,z1,MyNewTool\WObj:=Cara;
    ENDPROC
    PROC CicloDecoracion()
        ConveyorStop;
        ConveyorForward;
        WaitTime TiempoEntrada;
        ConveyorStop;
        WaitTime TiempoDeslizamiento;
        Set DO_01;
        RutinaDecoracion;
        Reset DO_01;
        Path_Home;
        ConveyorForward;
        WaitTime TiempoSalida;
        ConveyorStop;
        WaitTime TiempoDeslizamiento;
    ENDPROC
    PROC ConveyorForward()
        Reset BWD_Conveyor;
        WaitTime 0.2;
        Set FWD_Conveyor;
    ENDPROC
    PROC ConveyorBackward()
        Reset FWD_Conveyor;
        WaitTime 0.2;
        Set BWD_Conveyor;
    ENDPROC
    PROC ConveyorStop()
        Reset FWD_Conveyor;
        Reset BWD_Conveyor;
    ENDPROC

ENDMODULE
